(* IEC 61131-3 sources: plc-vscode/tests/st/non-utf8/rusty/tests/integration/data, 2 files *)

(* ---- encoding_utf_16.st ---- *)
PROGRAM a
(* Cömment *)
END_PROGRAM

(* ---- encoding_win.st ---- *)
PROGRAM a
(* Cömment *)
END_PROGRAM
